SUBAPPLICATION Uebung_149_AX (* Übung zu ETP senden (PGN 0x1EF00, 4000 Byte an das andere logiBUS) *)
  (* Standard: 61499-2; Description: Copyright (c) 2026 Meisterschulen am Ostbahnhof This program and the accompanying materials are made available under the terms of the Eclipse Public License 2.0 which is available at https://www.eclipse.org/legal/epl-2.0/ SPDX-License-Identifier: EPL-2.0 *)
  (* Version 1.0, 2026-11-17, Franz Höpfinger, Meisterschulen am Ostbahnhof, initial API and implementation and/or initial documentation *)
  PACKAGE Uebungen;
  IMPORT Uebungen::const::Uebung_140_149::Etp::LOGIBUS_ADD;
  IMPORT Uebungen::const::Uebung_140_149::Etp::LOGIBUS_FLT;
  IMPORT isobus::pgn::ISOUSERHOME_e::network;
  IMPORT isobus::pgn::ISO_CAN_NODE::NODE1;
  IMPORT isobus::pgn::const::PgnDef::PGN_PDU1_PropA2;
  IMPORT logiBUS::io::DI::logiBUS_DI::Input_I1;
  IMPORT logiBUS::io::DI::logiBUS_DI_Events::BUTTON_SINGLE_CLICK;
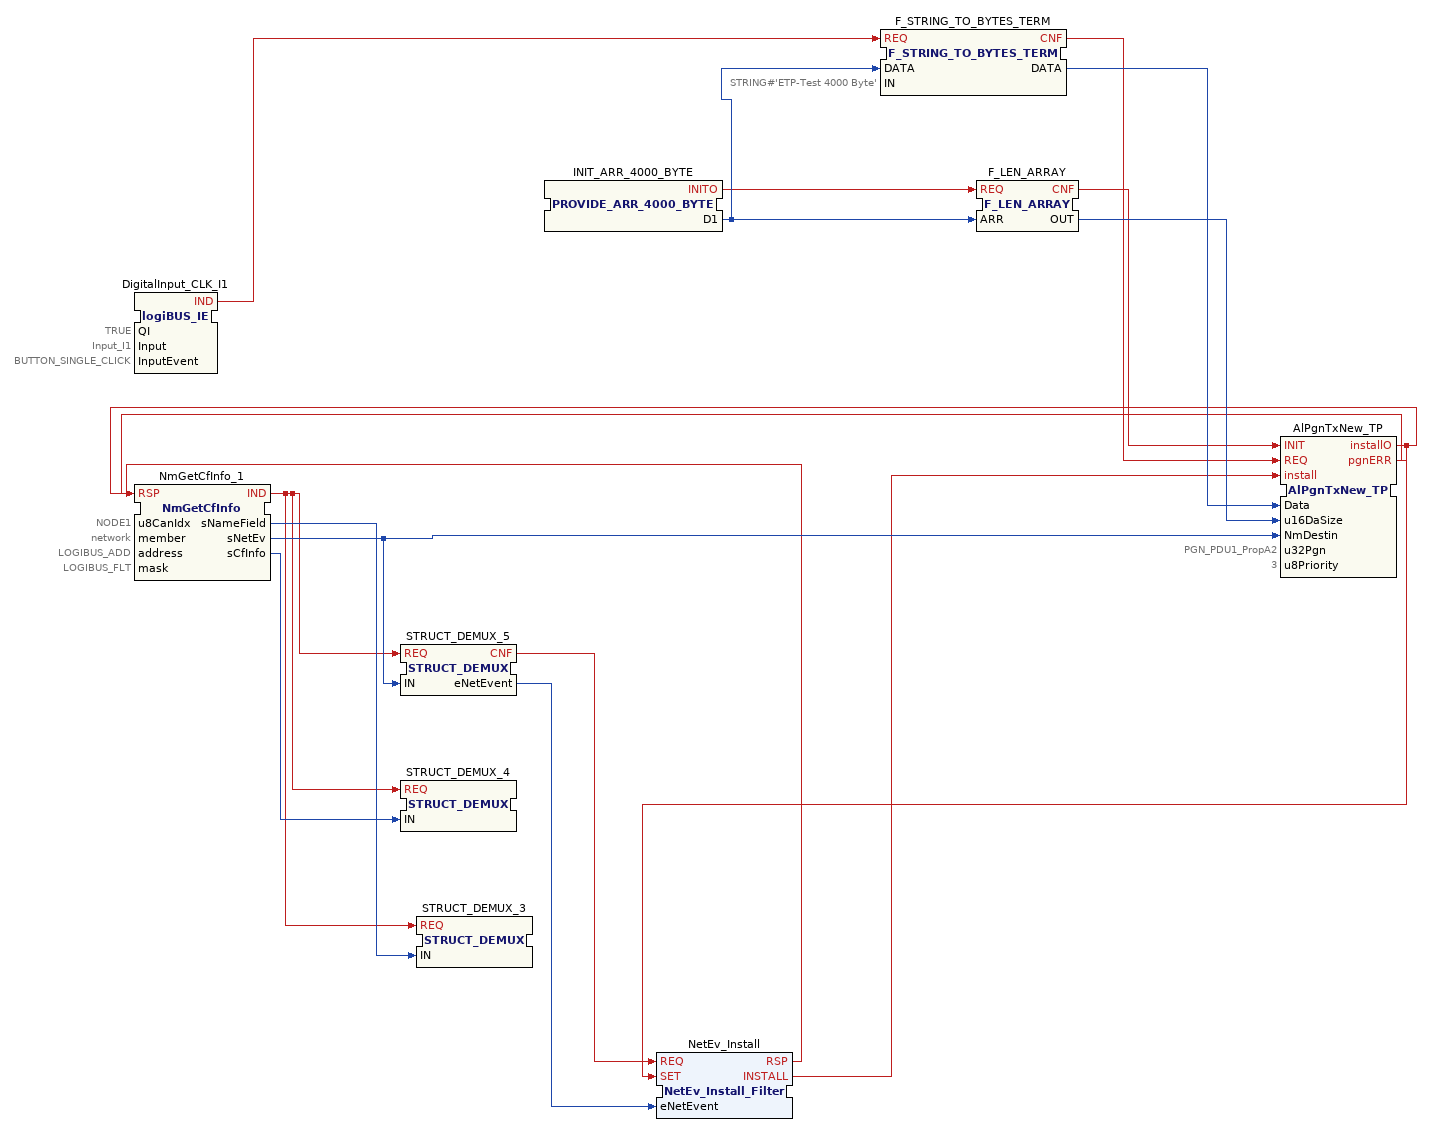
  (* ETP senden: PGN PropA2 0x1EF00, 4000 Byte an das andere logiBUS Mehr als 1785 Byte gehen per ETP (Extended Transport Protocol). Das geht nur an EINEN Empfänger, nicht global. Partner: NmGetCfInfo mit network + Filter LOGIBUS_ADD/LOGIBUS_FLT (Hersteller 1116, Funktion 128). I1 Klick sendet: Text ETP-Test 4000 Byte, dann 16#00, Rest 16#FF. Den Stack wählt TP oder ETP selbst. Gegenstück: Übung 149b (oder 149c mit zu kleinem Puffer). Nicht 0x1F000-0x1FFFF: das ist Fast Packet. Firmware ab LOGIBUS 24534469 auf BEIDEN Geräten. *)
  FBS
    STRUCT_DEMUX_3 : eclipse4diac::convert::STRUCT_DEMUX; {SET_ATTRIBUTE(StructuredType, isobus::pgn::NAMEFIELD_T)}
    NmGetCfInfo_1 : isobus::pgn::NmGetCfInfo(u8CanIdx := NODE1, member := network, address := LOGIBUS_ADD, mask := LOGIBUS_FLT);
    STRUCT_DEMUX_4 : eclipse4diac::convert::STRUCT_DEMUX; {SET_ATTRIBUTE(StructuredType, isobus::pgn::CF_INFO_T)}
    STRUCT_DEMUX_5 : eclipse4diac::convert::STRUCT_DEMUX; {SET_ATTRIBUTE(StructuredType, isobus::pgn::ISONETEVENT_T)}
    INIT_ARR_4000_BYTE : eclipse4diac::convert::providers::PROVIDE_ARR_4000_BYTE;
    F_LEN_ARRAY : eclipse4diac::utils::arrays::F_LEN_ARRAY;
    F_STRING_TO_BYTES_TERM : logiBUS::utils::dyn_arr::F_STRING_TO_BYTES_TERM(IN := STRING#'ETP-Test 4000 Byte');
    AlPgnTxNew_TP : isobus::pgn::tx::AlPgnTxNew_TP(u32Pgn := PGN_PDU1_PropA2, u8Priority := 3);
    DigitalInput_CLK_I1 : logiBUS::io::DI::logiBUS_IE(QI := TRUE, Input := Input_I1, InputEvent := BUTTON_SINGLE_CLICK);
  END_FBS
  SUBAPPS
    NetEv_Install : MyLib::sys::NetEv_Install_Filter;
  END_SUBAPPS
  EVENT_CONNECTIONS
    NmGetCfInfo_1.IND TO STRUCT_DEMUX_3.REQ;
    NmGetCfInfo_1.IND TO STRUCT_DEMUX_4.REQ;
    NmGetCfInfo_1.IND TO STRUCT_DEMUX_5.REQ;
    DigitalInput_CLK_I1.IND TO F_STRING_TO_BYTES_TERM.REQ;
    INIT_ARR_4000_BYTE.INITO TO F_LEN_ARRAY.REQ;
    F_LEN_ARRAY.CNF TO AlPgnTxNew_TP.INIT;
    F_STRING_TO_BYTES_TERM.CNF TO AlPgnTxNew_TP.REQ;
    AlPgnTxNew_TP.installO TO NmGetCfInfo_1.RSP;
    AlPgnTxNew_TP.pgnERR TO NmGetCfInfo_1.RSP;
    STRUCT_DEMUX_5.CNF TO NetEv_Install.REQ;
    NetEv_Install.RSP TO NmGetCfInfo_1.RSP;
    AlPgnTxNew_TP.installO TO NetEv_Install.SET;
    NetEv_Install.INSTALL TO AlPgnTxNew_TP.install;
  END_CONNECTIONS
  DATA_CONNECTIONS
    NmGetCfInfo_1.sNameField TO STRUCT_DEMUX_3.IN;
    NmGetCfInfo_1.sNetEv TO STRUCT_DEMUX_5.IN;
    NmGetCfInfo_1.sCfInfo TO STRUCT_DEMUX_4.IN;
    INIT_ARR_4000_BYTE.D1 TO F_LEN_ARRAY.ARR;
    INIT_ARR_4000_BYTE.D1 TO F_STRING_TO_BYTES_TERM.DATA;
    F_STRING_TO_BYTES_TERM.DATA TO AlPgnTxNew_TP.Data;
    F_LEN_ARRAY.OUT TO AlPgnTxNew_TP.u16DaSize;
    STRUCT_DEMUX_5.eNetEvent TO NetEv_Install.eNetEvent;
    NmGetCfInfo_1.sNetEv TO AlPgnTxNew_TP.NmDestin;
  END_CONNECTIONS
END_SUBAPPLICATION
